PROGRAM main
  VAR_INPUT
    Start_PB AT %IX0.0 : BOOL;
    Stop_PB AT %IX0.1 : BOOL;
    Sensor_1 AT %IX0.2 : BOOL;
    Sensor_2 AT %IX0.3 : BOOL;
  END_VAR
  VAR_OUTPUT
    Conveyor AT %QX0.0 : BOOL;
    Running_Lamp AT %QX0.1 : BOOL;
  END_VAR
  VAR
    Timer_1 : TON;
  END_VAR

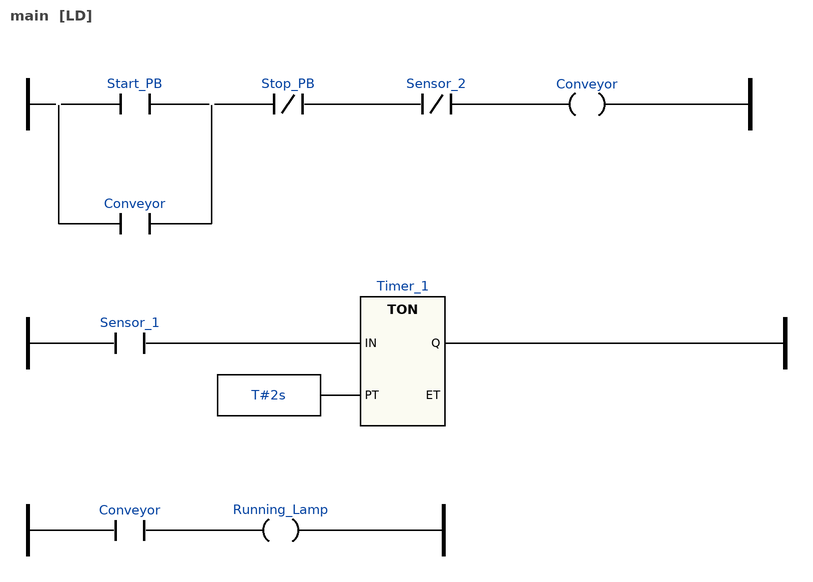
(* LD diagram, written out as Structured Text *)
Conveyor := (Start_PB OR Conveyor) AND NOT Stop_PB AND NOT Sensor_2;
Running_Lamp := Conveyor;
Timer_1(IN := Sensor_1, PT := T#2s);
END_PROGRAM
